(* IEC 61131-3 sources: plc-vscode/tests/st/test-ready/rusty/tests/integration/data/multi, 7 files *)

(* ---- concat_date.st ---- *)
{external}
FUNCTION CONCAT_DATE <T: ANY_INT> : DATE
VAR_INPUT
    year : T;
    month : T;
    day : T;
END_VAR
END_FUNCTION

(* ---- concat_date_prg1.st ---- *)
FUNCTION foo1 : LINT
    foo1 := CONCAT_DATE(INT#1, SINT#2, SINT#3);
END_FUNCTION

(* ---- concat_date_prg2.st ---- *)
FUNCTION foo2 : LINT
    foo2 := CONCAT_DATE(INT#4, SINT#5, SINT#6);
END_FUNCTION

(* ---- func.st ---- *)
FUNCTION main : INT
VAR_INPUT

END_VAR

VAR

END_VAR
mainProg();
main := mainProg.a;

END_FUNCTION

(* ---- enum1.st ---- *)
FUNCTION_BLOCK FOO
VAR
	foo_enum : (stop, go) := go;
END_VAR
END_FUNCTION_BLOCK

(* ---- enum2.st ---- *)
FUNCTION_BLOCK BAR
VAR
	bar_enum : (stop, go) := go;
END_VAR
END_FUNCTION_BLOCK

(* ---- prog.st ---- *)
PROGRAM mainProg
VAR
    a: DINT := 0;
END_VAR
a := 42;
END_PROGRAM
